// TIA Portal V20 export
// export: Created 2026-10-11T05:25:30.7219516Z, ExportSetting WithDefaults, DisplayName Totally Integrated Automation Portal, DisplayVersion V20, DisplayName TIA Portal Openness, DisplayVersion V20, DisplayName TIA Portal Teamcenter Gateway, DisplayVersion V20, DisplayName TIA Portal Version Control Interface, DisplayVersion V20, DisplayName SINAMICS Startdrive Advanced, DisplayVersion V20 SP1 Update 2, DisplayName SINAMICS Startdrive G110M, G120, G120C, G120D, G120P, G115D, DisplayVersion V20 SP1 Update 2, DisplayName SINAMICS Startdrive G130, G150, S120, S150, SINAMICS MV, G220, S200, S210, DisplayVersion V20 SP1 Update 2, DisplayName STEP 7 Professional, DisplayVersion V20, DisplayName STEP 7 Safety, DisplayVersion V20, DisplayName WinCC Basic/Comfort/Advanced, DisplayVersion V20, DisplayName WinCC Professional, DisplayVersion V20, DisplayName WinCC Unified, DisplayVersion V20
FUNCTION "FRK_PartProcessed" : Bool   // FC40, SCL
{ S7_Optimized_Access := 'TRUE' }
VERSION : 0.1
// stored: AutoNumber true, IsIECCheckEnabled false, SetENOAutomatically false, UDAEnableTagReadback false
   VAR_INPUT
      Verdict : DInt;
      Reason : DInt;
   END_VAR
   VAR_IN_OUT
      Core : "FRK_Core";
      Unit : "FRK_Unit";
      Status : "ST_ModuleStatus";
      Part : "ST_PartContext";
      History : Array[1..16] of "ST_Diagnostic";
      Head : Int;
   END_VAR
   VAR_TEMP
      Index : DInt;
      Stamp : DTL;
      ResultCode : Int;
   END_VAR
BEGIN

   #FRK_PartProcessed := FALSE;
   #Index := #Unit.CarrierIndex;
   IF #Index = 0 OR NOT #Part.Present THEN
       RETURN;
   END_IF;
   IF #Verdict < 1 OR #Verdict > 3 OR (#Verdict = 2 AND #Reason = 0) THEN
       "FRK_Fault"(Core := #Core,
                   Status := #Status,
                   ReasonCode := 2023,
                   Description := WSTRING#'std.error.nokReasonRequired');
       RETURN;
   END_IF;
   IF #Index < 1 OR #Index > 32 THEN
       "FRK_Fault"(Core := #Core,
                   Status := #Status,
                   ReasonCode := 2021,
                   Description := WSTRING#'std.error.partCarrierWriteFailed');
       RETURN;
   END_IF;
   IF NOT "FRK_Carriers".Slots[#Index].Enabled THEN
       "FRK_Fault"(Core := #Core,
                   Status := #Status,
                   ReasonCode := 2021,
                   Description := WSTRING#'std.error.partCarrierWriteFailed');
       RETURN;
   END_IF;
   IF #Part.Uid <> "FRK_Carriers".Slots[#Index].Context.Uid THEN
       "FRK_Fault"(Core := #Core,
                   Status := #Status,
                   ReasonCode := 2022,
                   Description := WSTRING#'std.error.partCarrierReadFailed');
       RETURN;
   END_IF;
   #Part.Result.Verdict := #Verdict;
   #Part.Result.ReasonCode := #Reason;
   #Part.Result.StationPath := STRING_TO_WSTRING(#Status.Name);
   #Part.Result.TimeSynchronized := FALSE;
   #ResultCode := RD_SYS_T(OUT => #Stamp);
   IF #ResultCode = 0 THEN
       #Part.Result.Stamp := DTL_TO_LDT(#Stamp);
   END_IF;
   "FRK_Carriers".Slots[#Index].Written := #Part;
   IF "FRK_Carriers".Slots[#Index].Writes < UDINT#4294967295 THEN
       "FRK_Carriers".Slots[#Index].Writes := "FRK_Carriers".Slots[#Index].Writes + 1;
   END_IF;
   CASE #Verdict OF
       1:
           IF #Unit.Good < UDINT#4294967295 THEN
               #Unit.Good := #Unit.Good + 1;
           END_IF;
       2:
           IF #Unit.Nok < UDINT#4294967295 THEN
               #Unit.Nok := #Unit.Nok + 1;
           END_IF;
           #Unit.NokReason := #Reason;
       3:
           IF #Unit.Rework < UDINT#4294967295 THEN
               #Unit.Rework := #Unit.Rework + 1;
           END_IF;
       ELSE
           RETURN;
   END_CASE;
   // The provider result is written before publishing EVENT_PART_PROCESSED.
   "FRK_PartEvent"(History := #History,
                   Head := #Head,
                   Reason := 2026,
                   Uid := #Part.Uid,
                   SourcePath := #Status.Name);
   #Part.Present := FALSE;
   #FRK_PartProcessed := TRUE;
END_FUNCTION
